                                           //Is the data in the tcp receive buffer to be analyzed bigger than 1 byte
                                           IF (#statReceive.trcvFct.dataLengthRest > 1) THEN
                                               //Yes --> get the telegram type in the 2nd byte
                                               #statReceive.tempTelegram.telegramType := #statReceive.trcvFct.data[#statReceive.trcvFct.dataOffset + 1];
                                           ELSE
                                               //No --> just one byte
                                               #statCopyNBytes := 1;
                                               #statReceive.tempTelegram.telegramType := 0;
                                           END_IF;

                                       ELSE
                                           //Already data in the temp. LCom header
                                           IF (#statReceive.tempTelegram.index = 1) THEN
                                               //Get the telegram type in the 1st byte
                                               #statReceive.tempTelegram.telegramType := #statReceive.trcvFct.data[#statReceive.trcvFct.dataOffset];
                                           ELSE
                                               //Get the telegram type in the 2nd byte
                                               #statReceive.tempTelegram.telegramType := #statReceive.trcvFct.data[#statReceive.trcvFct.dataOffset + 1];
                                           END_IF;
                                       END_IF;


                                       //---------------------------------------------------------------------
                                       //Build temp LCom header, if the telegram type is known
                                       //---------------------------------------------------------------------
                                       //Check if the telegram type is known
                                       IF (#statReceive.tempTelegram.telegramType > 0) THEN

                                           //Yes -->  telegram type is known
                                           CASE (#statReceive.tempTelegram.telegramType) OF
                                               1..3://Config telegram type 1,2,3
                                                   //LCom V2 (24 byte)
                                                   IF (#statReceive.tempTelegram.LComVersion = #HEADER_V2) THEN
                                                       IF ((24 - #statReceive.tempTelegram.index) < #statReceive.trcvFct.dataLengthRest) THEN
                                                           #statCopyNBytes := 24 - #statReceive.tempTelegram.index;
                                                       ELSE
                                                           #statCopyNBytes := #statReceive.trcvFct.dataLengthRest;
                                                       END_IF;
                                                   ELSE
                                                       //LCom V1 (16 byte)
                                                       IF ((16 - #statReceive.tempTelegram.index) < #statReceive.trcvFct.dataLengthRest) THEN
                                                           #statCopyNBytes := 16 - #statReceive.tempTelegram.index;
                                                       ELSE
                                                           #statCopyNBytes := #statReceive.trcvFct.dataLengthRest;
                                                       END_IF;
                                                   END_IF;
                                               5://Clock synchronization telegram type 5
                                                   //LCom V1 and V2 (10 byte)
                                                   IF ((10 - #statReceive.tempTelegram.index) < #statReceive.trcvFct.dataLengthRest) THEN
                                                       #statCopyNBytes := 10 - #statReceive.tempTelegram.index;
                                                   ELSE
                                                       #statCopyNBytes := #statReceive.trcvFct.dataLengthRest;
                                                   END_IF;
                                               10://Data telegram type 10
                                                   //LCom V2 (20 byte)
                                                   IF (#statReceive.tempTelegram.LComVersion = #HEADER_V2) THEN
                                                       IF ((20 - #statReceive.tempTelegram.index) < #statReceive.trcvFct.dataLengthRest) THEN
                                                           #statCopyNBytes := 20 - #statReceive.tempTelegram.index;
                                                       ELSE
                                                           #statCopyNBytes := #statReceive.trcvFct.dataLengthRest;
                                                       END_IF;
                                                   ELSE
                                                       //LCom V1 (12 byte)
                                                       IF ((12 - #statReceive.tempTelegram.index) < #statReceive.trcvFct.dataLengthRest) THEN
                                                           #statCopyNBytes := 12 - #statReceive.tempTelegram.index;
                                                       ELSE
                                                           #statCopyNBytes := #statReceive.trcvFct.dataLengthRest;
                                                       END_IF;
                                                   END_IF;
                                               20://Close connection telegram type 20
                                                   //LCom V1 (2 byte)
                                                   IF ((2 - #statReceive.tempTelegram.index) < #statReceive.trcvFct.dataLengthRest) THEN
                                                       #statCopyNBytes := 2 - #statReceive.tempTelegram.index;
                                                   ELSE
                                                       #statCopyNBytes := #statReceive.trcvFct.dataLengthRest;
                                                   END_IF;
                                               ELSE
                                                   //Write diagnostics
                                                   #statDiag.bufferIndex := #statDiag.bufferIndex + 1;
                                                   #statDiag.buffer[#statDiag.bufferIndex].status := #ERR_WRONG_TELEGRAM_ID;
                                                   #statDiag.buffer[#statDiag.bufferIndex].subFunctionErrorID := 16#0000;
                                                   #statDiag.buffer[#statDiag.bufferIndex].additionalValue1 := #statReceive.tempTelegram.telegramType;
                                                   #statDiag.buffer[#statDiag.bufferIndex].additionalValue2 := 0.0;
                                                   #statDiag.buffer[#statDiag.bufferIndex].additionalValue3 := 0.0;
                                                   #statDiag.buffer[#statDiag.bufferIndex].additionalValue4 := T#0ms;

                                                   #statState.connection := #CLOSE_CONNECTION;
                                                   GOTO diag;
                                           END_CASE;
                                       ELSE
                                           ;//No --> telegram type is zero
                                       END_IF;

                                       //Copy data into the temp. LCom header
                                       #statRet := MOVE_BLK_VARIANT(SRC := #statReceive.trcvFct.data, COUNT := #statCopyNBytes, SRC_INDEX := UDINT_TO_DINT(#statReceive.trcvFct.dataOffset), DEST_INDEX := #statReceive.tempTelegram.index, DEST => #statReceive.tempTelegram.data);
                                       //Calculate index in the temp. LCom header buffer
                                       #statReceive.tempTelegram.index := #statReceive.tempTelegram.index + UDINT_TO_USINT(#statCopyNBytes);
                                       //Calculate offset in the tcp receive buffer
                                       #statReceive.trcvFct.dataOffset := #statReceive.trcvFct.dataOffset + #statCopyNBytes;

                                       //Is local LCom version equal to partner LCom version ?
                                       IF (#statActualLocalLComVersion <> #statReceive.tempTelegram.LComVersion) THEN
                                           #statConnectAttempts := #statConnectAttempts + 1;
                                           //Write diagnostics
                                           #statDiag.bufferIndex := #statDiag.bufferIndex + 1;
                                           #statDiag.buffer[#statDiag.bufferIndex].status := #ERR_WRONG_HEADER;
                                           #statDiag.buffer[#statDiag.bufferIndex].subFunctionErrorID := 16#0000;
                                           #statDiag.buffer[#statDiag.bufferIndex].additionalValue1 := #statReceive.tempTelegram.LComVersion;
                                           #statDiag.buffer[#statDiag.bufferIndex].additionalValue2 := #statActualLocalLComVersion;
                                           #statDiag.buffer[#statDiag.bufferIndex].additionalValue3 := 0.0;
                                           #statDiag.buffer[#statDiag.bufferIndex].additionalValue4 := T#0ms;

                                           #statState.connection := #CLOSE_CONNECTION;
                                           GOTO diag;
                                       ELSE
                                           ;//local LCom version and partner LCom versions are equal
                                           #diagnostics.statistics.activeLComVersion := #statActualLocalLComVersion;
                                       END_IF;
                                   END_IF;//End: There is data expected without LCom header

                                   //---------------------------------------------------------------------
                                   //Interpret temp LCom header
                                   //---------------------------------------------------------------------
                                   IF (((#statReceive.tempTelegram.LComVersion = #HEADER_V1)//LCom V1
                                       AND//1,2,3 = 16 Byte
                                       ((#statReceive.tempTelegram.telegramType <= 3 AND #statReceive.tempTelegram.index = 16)
                                       OR//5 = 10 Byte
                                       (#statReceive.tempTelegram.telegramType = 5 AND #statReceive.tempTelegram.index = 10)
                                       OR//10 = 12 Byte
                                       (#statReceive.tempTelegram.telegramType = 10 AND #statReceive.tempTelegram.index = 12)
                                       OR//20 = 2 Byte
                                       (#statReceive.tempTelegram.telegramType = 20 AND #statReceive.tempTelegram.index = 2)))
                                       OR
                                       ((#statReceive.tempTelegram.LComVersion = #HEADER_V2)//LCom V2
                                       AND//1,2,3 = 24 Byte
                                       ((#statReceive.tempTelegram.telegramType <= 3 AND #statReceive.tempTelegram.index = 24)
                                       OR//5 = 10 Byte
                                       (#statReceive.tempTelegram.telegramType = 5 AND #statReceive.tempTelegram.index = 10)
                                       OR//10 = 20 Byte
                                       (#statReceive.tempTelegram.telegramType = 10 AND #statReceive.tempTelegram.index = 20)))
                                       OR
                                       (#statState.comReceiver = #DATA_EXPECTED))
                                   THEN

                                       CASE #statReceive.tempTelegram.telegramType OF

                                           10://Telegram type 10

                                               //Data expected without LCom header ?
                                               IF (#statState.comReceiver = #DATA_EXPECTED) THEN
                                                   //Yes --> LCom header from data telegram is already interpreted
                                                   //#receive.dataTelegram.messageOffset and #receive.dataTelegram.acPackageLength is known
                                                   //Calculate the bytes which have to be copied into FB.receiveData
                                                   IF (#statReceive.userData.offset + #statReceive.trcvFct.dataLengthRest) > (#statReceive.dataTelegram.messageOffset + #statReceive.dataTelegram.actPackageLength) THEN
                                                       //Copy just the missing bytes from the actual LCom package
                                                       #statCopyNBytes := ((#statReceive.dataTelegram.messageOffset + #statReceive.dataTelegram.actPackageLength) - #statReceive.userData.offset);
                                                   ELSE
                                                       //Copy all bytes which are still in the tcp receive buffer
                                                       #statCopyNBytes := #statReceive.trcvFct.dataLengthRest;
                                                   END_IF;
                                                   //Set SEND acknowledge message offset
                                                   #statSend.dataTelegram.ackMessageOffset := #statSend.dataTelegram.ackMessageOffset + #statCopyNBytes;
                                               ELSE
                                                   //Reset index, so a new temp. LCom header can be build
                                                   #statReceive.tempTelegram.index := 0;
                                                   #statReceive.numberOfLComHeader := #statReceive.numberOfLComHeader + 1;

                                                   //LComVersion
                                                   #statReceive.dataTelegram.LComVersion := #statReceive.tempTelegram.data[0];
                                                   //Telegram type
                                                   #statReceive.dataTelegram.telegramType := #statReceive.tempTelegram.data[1];
                                                   //Message counter
                                                   #statReceive.dataTelegram.messageCounter := #statReceive.tempTelegram.data[2];
                                                   //Acknowledge message counter
                                                   #statReceive.dataTelegram.ackMessageCounter := #statReceive.tempTelegram.data[3];

                                                   //LCom V2
                                                   IF (#statActualLocalLComVersion = #HEADER_V2) THEN
                                                       //Get tem. total message length
                                                       #tempDWord.%B3 := #statReceive.tempTelegram.data[16];
                                                       #tempDWord.%B2 := #statReceive.tempTelegram.data[17];
                                                       #tempDWord.%B1 := #statReceive.tempTelegram.data[18];
                                                       #tempDWord.%B0 := #statReceive.tempTelegram.data[19];

                                                       //Acknowledge message offset
                                                       #statReceive.dataTelegram.ackMessageOffset.%B3 := #statReceive.tempTelegram.data[8];
                                                       #statReceive.dataTelegram.ackMessageOffset.%B2 := #statReceive.tempTelegram.data[9];
                                                       #statReceive.dataTelegram.ackMessageOffset.%B1 := #statReceive.tempTelegram.data[10];
                                                       #statReceive.dataTelegram.ackMessageOffset.%B0 := #statReceive.tempTelegram.data[11];

                                                       //Is it an acknowledge telegram ?
                                                       IF (#tempDWord = 16#0000) THEN
                                                           //Acknowledge telegram
                                                           #statState.comReceiver := #ACK_TELEGRAM;
                                                       ELSE
                                                           //Is no acknowledge telegram
                                                           //Message offset
                                                           #statReceive.dataTelegram.messageOffset.%B3 := #statReceive.tempTelegram.data[4];
                                                           #statReceive.dataTelegram.messageOffset.%B2 := #statReceive.tempTelegram.data[5];
                                                           #statReceive.dataTelegram.messageOffset.%B1 := #statReceive.tempTelegram.data[6];
                                                           #statReceive.dataTelegram.messageOffset.%B0 := #statReceive.tempTelegram.data[7];
                                                           //Actual package length
                                                           #statReceive.dataTelegram.actPackageLength.%B3 := #statReceive.tempTelegram.data[12];
                                                           #statReceive.dataTelegram.actPackageLength.%B2 := #statReceive.tempTelegram.data[13];
                                                           #statReceive.dataTelegram.actPackageLength.%B1 := #statReceive.tempTelegram.data[14];
                                                           #statReceive.dataTelegram.actPackageLength.%B0 := #statReceive.tempTelegram.data[15];
                                                           //Total message length
                                                           #statReceive.dataTelegram.totalMessageLength := #tempDWord;
                                                       END_IF;
                                                   ELSE
                                                       //LCom V1
                                                       //Get temp. total message length
                                                       #tempDWord.%B1 := #statReceive.tempTelegram.data[10];
                                                       #tempDWord.%B0 := #statReceive.tempTelegram.data[11];

                                                       //Acknowledge message offset
                                                       #statReceive.dataTelegram.ackMessageOffset.%B1 := #statReceive.tempTelegram.data[6];
                                                       #statReceive.dataTelegram.ackMessageOffset.%B0 := #statReceive.tempTelegram.data[7];

                                                       //Is it an acknowledge telegram ?
                                                       IF (#tempDWord = 16#0000) THEN
                                                           //Acknowledge telegram
                                                           #statState.comReceiver := #ACK_TELEGRAM;
                                                       ELSE
                                                           //Is no acknowledge telegram
                                                           //Message offset
                                                           #statReceive.dataTelegram.messageOffset.%B1 := #statReceive.tempTelegram.data[4];
                                                           #statReceive.dataTelegram.messageOffset.%B0 := #statReceive.tempTelegram.data[5];
                                                           //Actual package length
                                                           #statReceive.dataTelegram.actPackageLength.%B1 := #statReceive.tempTelegram.data[8];
                                                           #statReceive.dataTelegram.actPackageLength.%B0 := #statReceive.tempTelegram.data[9];
                                                           //Total message length
                                                           #statReceive.dataTelegram.totalMessageLength := #tempDWord;
                                                       END_IF;
                                                   END_IF;

                                                   //Set SEND acknowledge message offset
                                                   #statSend.dataTelegram.ackMessageCounter := #statReceive.dataTelegram.messageCounter;

                                                   //Check if the LCom package, which was sent before is acknowledged ?
                                                   IF ((#statSend.numberOfLComPackage = 1)//One package was sent
                                                       AND
                                                       ((#statSend.expectedAck.package1.offset = #statReceive.dataTelegram.ackMessageOffset)
                                                       AND
                                                       (#statSend.dataTelegram.messageCounter = #statReceive.dataTelegram.ackMessageCounter)))
                                                   THEN
                                                       //Acknowledgement for the package x.1
                                                       #statSend.numberOfLComPackage := 0;
                                                       //Stop acknowledge timer for the 1st package
                                                       #instExpectedAckPackage1(IN := FALSE,
                                                                                PT := #diagnostics.localConfig.sender.ackTimeout);
                                                   ELSIF ((#statSend.dataTelegram.messageCounter = #statReceive.dataTelegram.ackMessageCounter)
                                                       OR
                                                       (#statSend.dataTelegram.messageCounter - 1 = #statReceive.dataTelegram.ackMessageCounter)
                                                       OR
                                                       (#diagnostics.statistics.maxMsgSendingTime = T#0ms))//Workaround: S7 Controller does not start with correct ack. message counter
                                                   THEN
                                                       ;
                                                   ELSE
                                                       //Write diagnostics
                                                       #statDiag.bufferIndex := #statDiag.bufferIndex + 1;
                                                       #statDiag.buffer[#statDiag.bufferIndex].status := #ERR_ACK_MESSAGE_NUMBER;
                                                       #statDiag.buffer[#statDiag.bufferIndex].subFunctionErrorID := 16#0000;
                                                       #statDiag.buffer[#statDiag.bufferIndex].additionalValue1 := #statReceive.dataTelegram.messageCounter;
                                                       #statDiag.buffer[#statDiag.bufferIndex].additionalValue2 := #statSend.dataTelegram.messageCounter;
                                                       #statDiag.buffer[#statDiag.bufferIndex].additionalValue3 := 0.0;
                                                       #statDiag.buffer[#statDiag.bufferIndex].additionalValue4 := T#0ms;

                                                       #statState.connection := #CLOSE_CONNECTION;
                                                       GOTO diag;
                                                   END_IF;


                                                   //Is the 1st LCom package received and nothing is copied into FB.receiveData so far ?
                                                   IF ((#statReceive.userData.totalLength = 0)
                                                       AND
                                                       (#statReceive.dataTelegram.messageOffset = 0)
                                                       AND
                                                       (#statState.comReceiver <> #ACK_TELEGRAM))
                                                   THEN
                                                       //Store the 1st received telegram with the total receive length
                                                       #statReceive.userData.totalLength := #statReceive.dataTelegram.totalMessageLength;
                                                       //Reset the acknowledged message offset
                                                       #statSend.dataTelegram.ackMessageOffset := 0;

                                                       //Start message receiving timer
                                                       #instMsgReceivingTimer(IN := TRUE,
                                                                              PT := T#+24d20h31m23s647ms);
                                                   ELSE
                                                       ;//In receiving process or acknowledge telegram
                                                   END_IF;

                                                   //Is the data telegram a acknowledge telegram ?
                                                   IF (#statState.comReceiver = #ACK_TELEGRAM)
                                                   THEN
                                                       //Yes --> Acknowledge telegram, no bytes have to be copied
                                                       #statCopyNBytes := 0;
                                                   ELSIF ((#diagnostics.statistics.activeLComVersion = #HEADER_V1)
                                                       AND
                                                       ((#statReceive.userData.offset + (#statReceive.trcvFct.dataLengthRest - 12)) > (#statReceive.dataTelegram.messageOffset + #statReceive.dataTelegram.actPackageLength)))
                                                   THEN//No --> The data to be analyzed in the tcp receive buffer is bigger than the complete message

                                                       //Do not copy all data from the tcp receive buffer, only the rest data from the LCom package
                                                       #statCopyNBytes := ((#statReceive.dataTelegram.messageOffset + #statReceive.dataTelegram.actPackageLength) - #statReceive.userData.offset);
                                                       //Calculate acknowledge message offset which has to be sent to the partner
                                                       #statSend.dataTelegram.ackMessageOffset := #statSend.dataTelegram.ackMessageOffset + #statCopyNBytes;
                                                   ELSIF ((#diagnostics.statistics.activeLComVersion = #HEADER_V2)
                                                       AND
                                                       ((#statReceive.userData.offset + (#statReceive.trcvFct.dataLengthRest - 24)) > (#statReceive.dataTelegram.messageOffset + #statReceive.dataTelegram.actPackageLength)))
                                                   THEN//No --> The data to be analyzed in the tcp receive buffer is bigger than the complete message

                                                       //Copy not all data from the tcp receive buffer, only the rest data from the LCom package
                                                       #statCopyNBytes := ((#statReceive.dataTelegram.messageOffset + #statReceive.dataTelegram.actPackageLength) - #statReceive.userData.offset);
                                                       //Calculate acknowledge message offset which have to be sent to the partner
                                                       #statSend.dataTelegram.ackMessageOffset := #statSend.dataTelegram.ackMessageOffset + #statCopyNBytes;
                                                   ELSE
                                                       //Copy just the rest of data from the tcp receive buffer
                                                       IF #diagnostics.statistics.activeLComVersion = #HEADER_V1 THEN
                                                           #statCopyNBytes := #statReceive.trcvFct.dataLengthRest - 12;
                                                       ELSE
                                                           #statCopyNBytes := #statReceive.trcvFct.dataLengthRest - 20;
                                                       END_IF;
                                                       //Calculate acknowledge message offset which have to be sent to the partner
                                                       #statSend.dataTelegram.ackMessageOffset := #statSend.dataTelegram.ackMessageOffset + #statCopyNBytes;
                                                   END_IF;

                                               END_IF;

                                               //Copy data to FB.receiveBuffer
                                               #statRet := MOVE_BLK_VARIANT(SRC := #statReceive.trcvFct.data, COUNT := #statCopyNBytes, SRC_INDEX := UDINT_TO_DINT(#statReceive.trcvFct.dataOffset), DEST_INDEX := UDINT_TO_DINT(#statReceive.userData.offset), DEST => #receiveBuffer);
                                               //Calculate offset in the FB.#receiveBuffer
                                               #statReceive.userData.offset := #statReceive.userData.offset + #statCopyNBytes;
                                               //Calculate offset in the tcp receive buffer
                                               #statReceive.trcvFct.dataOffset := #statReceive.trcvFct.dataOffset + #statCopyNBytes;

                                               //---------------------------------------------------------------------
                                               //Is complete LCom message acknowledged which was sent ?
                                               //---------------------------------------------------------------------
                                               IF ((#statSend.userData.offset = #statReceive.dataTelegram.ackMessageOffset)
                                                   AND
                                                   (#statReceive.dataTelegram.ackMessageCounter = #statSend.dataTelegram.messageCounter)
                                                   AND
                                                   #statState.comSender = #SEND_NO_DATA)
                                               THEN
                                                   //Yes --> Complete LCom message is acknowledged
                                                   #sending := #statSending := FALSE;

                                                   //Statistic --> Increase number of sent user messages
                                                   #diagnostics.statistics.numberOfSentMessages := #diagnostics.statistics.numberOfSentMessages + 1;

                                                   //Get message sending time [ms]
                                                   #instMsgSendingTimer(IN := TRUE,
                                                                        PT := T#+24d20h31m23s647ms);

                                                   //Statistic --> Compare max. message sending time
                                                   IF (#instMsgSendingTimer.ET > #diagnostics.statistics.maxMsgSendingTime) THEN
                                                       #diagnostics.statistics.maxMsgSendingTime := #instMsgSendingTimer.ET;
                                                   ELSE
                                                       ;//Actual sending time is smaller
                                                   END_IF;

                                                   //Statistic --> Calculate average of message sending time [ms)]
                                                   #diagnostics.statistics.avgMsgSendingTime := (((#diagnostics.statistics.avgMsgSendingTime * 19) + UDINT_TO_REAL((TIME_TO_UDINT(#instMsgSendingTimer.ET)))) / 20);

                                                   //Stop message sending timer
                                                   #instMsgSendingTimer(IN := FALSE,
                                                                        PT := T#+24d20h31m23s647ms);

                                                   //Initialize values, for next send request
                                                   #statSend.userData.offset := 0;
                                                   #statSend.dataTelegram.messageOffset := 0;
                                                   #statSend.dataTelegram.totalMessageLength := 0;
                                               ELSE
                                                   ;//Complete LCom message is not acknowledged yet
                                               END_IF;//End: Is complete Lcom message acknowledged, which was sent ?


                                               //---------------------------------------------------------------------
                                               //Build acknowledge telegram
                                               //---------------------------------------------------------------------

                                               //Assume always that an LCom package is expected
                                               #statState.comReceiver := #EXPECTED;

                                               //---------------------------------------------------------------------
                                               //Has the complete LCom package been received (1 Byte ... 4 Kilobyte) ?
                                               //---------------------------------------------------------------------
                                               IF (#statReceive.userData.offset = 0) THEN
                                                   ;//Do nothing
                                               ELSIF (#statReceive.userData.offset = (#statReceive.dataTelegram.messageOffset + #statReceive.dataTelegram.actPackageLength))
                                               THEN//Yes --> Complete LCom package has been received (1 Byte ... 4k Byte)

                                                   //Still in sending process and LCom package sent is not acknowledged yet ?
                                                   //Select LCom V1 or V2; now one LCom package is sent and must be acknowledged
                                                   IF ((#statSending = TRUE)
                                                       AND
                                                       (#statSend.numberOfLComPackage = 0)
                                                       AND
                                                       ((#statActualLocalLComVersion = #HEADER_V1)
                                                       OR
                                                       (#statActualLocalLComVersion = #HEADER_V2)))
                                                   THEN
                                                       ;//Build no acknowledge telegram 10
                                                   ELSE
                                                       //Build acknowledge telegram 10
                                                       #statSend.tsendFct.data[#statSend.tsendFct.dataOffset] := #statSend.dataTelegram.LComVersion;
                                                       #statSend.tsendFct.data[#statSend.tsendFct.dataOffset + 1] := #statSend.dataTelegram.telegramType;
                                                       #statSend.tsendFct.data[#statSend.tsendFct.dataOffset + 2] := #statSend.dataTelegram.messageCounter;
                                                       #statSend.tsendFct.data[#statSend.tsendFct.dataOffset + 3] := #statSend.dataTelegram.ackMessageCounter;
                                                       //Message offset
                                                       #statSend.tsendFct.data[#statSend.tsendFct.dataOffset + 4] := 16#00;
                                                       #statSend.tsendFct.data[#statSend.tsendFct.dataOffset + 5] := 16#00;
                                                       #statSend.tsendFct.data[#statSend.tsendFct.dataOffset + 6] := 16#00;
                                                       #statSend.tsendFct.data[#statSend.tsendFct.dataOffset + 7] := 16#00;
                                                       //Acknowledge message offset
                                                       #statSend.tsendFct.data[#statSend.tsendFct.dataOffset + 8] := #statSend.dataTelegram.ackMessageOffset.%B3;
                                                       #statSend.tsendFct.data[#statSend.tsendFct.dataOffset + 9] := #statSend.dataTelegram.ackMessageOffset.%B2;
                                                       #statSend.tsendFct.data[#statSend.tsendFct.dataOffset + 10] := #statSend.dataTelegram.ackMessageOffset.%B1;
                                                       #statSend.tsendFct.data[#statSend.tsendFct.dataOffset + 11] := #statSend.dataTelegram.ackMessageOffset.%B0;
                                                       //Actual package length
                                                       #statSend.tsendFct.data[#statSend.tsendFct.dataOffset + 12] := 16#00;
                                                       #statSend.tsendFct.data[#statSend.tsendFct.dataOffset + 13] := 16#00;
                                                       #statSend.tsendFct.data[#statSend.tsendFct.dataOffset + 14] := 16#00;
                                                       #statSend.tsendFct.data[#statSend.tsendFct.dataOffset + 15] := 16#00;
                                                       //Total message length
                                                       #statSend.tsendFct.data[#statSend.tsendFct.dataOffset + 16] := 16#00;
                                                       #statSend.tsendFct.data[#statSend.tsendFct.dataOffset + 17] := 16#00;
                                                       #statSend.tsendFct.data[#statSend.tsendFct.dataOffset + 18] := 16#00;
                                                       #statSend.tsendFct.data[#statSend.tsendFct.dataOffset + 19] := 16#00;

                                                       //LCom V2
                                                       IF (#statActualLocalLComVersion = #HEADER_V2) THEN
                                                           //Calculate offset in the tcp send buffer
                                                           #statSend.tsendFct.dataOffset := #statSend.tsendFct.dataOffset + 20;
                                                       ELSE
                                                           //LCom V1
                                                           //Acknowledge message offset
                                                           #statSend.tsendFct.data[#statSend.tsendFct.dataOffset + 6] := #statSend.dataTelegram.ackMessageOffset.%B1;
                                                           #statSend.tsendFct.data[#statSend.tsendFct.dataOffset + 7] := #statSend.dataTelegram.ackMessageOffset.%B0;
                                                           //Actual package length
                                                           #statSend.tsendFct.data[#statSend.tsendFct.dataOffset + 8] := 16#00;
                                                           #statSend.tsendFct.data[#statSend.tsendFct.dataOffset + 9] := 16#00;
                                                           //Total message length
                                                           #statSend.tsendFct.data[#statSend.tsendFct.dataOffset + 10] := 16#00;
                                                           #statSend.tsendFct.data[#statSend.tsendFct.dataOffset + 11] := 16#00;
                                                           //Calculate offset in the tcp send buffer
                                                           #statSend.tsendFct.dataOffset := #statSend.tsendFct.dataOffset + 12;
                                                       END_IF;
                                                       //Set sender state
                                                       #statState.sender := #SEND_CONFIG;
                                                   END_IF;


                                                   //---------------------------------------------------------------------
                                                   //Is the complete LCom message received (1 Byte ... 4 Gigabyte) ?
                                                   //---------------------------------------------------------------------
                                                   IF (#statReceive.userData.offset = #statReceive.dataTelegram.totalMessageLength) THEN
                                                       //Yes --> Set FB outputs
                                                       #dataReceived := #statDataReceived := TRUE;
                                                       #receivedDataLength := #statReceive.dataTelegram.totalMessageLength;
                                                       //Initialize values, for next receive request
                                                       #statReceive.userData.totalLength := 0;
                                                       #statReceive.userData.offset := 0;

                                                       //Statistic --> Increase number of received user messages
                                                       #diagnostics.statistics.numberOfReceivedMessages := #diagnostics.statistics.numberOfReceivedMessages + 1;

                                                       //Get message receiving time [ms]
                                                       #instMsgReceivingTimer(IN := TRUE,
                                                                              PT := T#+24d20h31m23s647ms);

                                                       //Statistic --> Compare max. message receiving time
                                                       IF (#instMsgReceivingTimer.ET > #diagnostics.statistics.maxMsgReceivingTime) THEN
                                                           #diagnostics.statistics.maxMsgReceivingTime := #instMsgReceivingTimer.ET;
                                                       ELSE
                                                           ;//Actual receiving time is smaller
                                                       END_IF;

                                                       //Statistic --> Calculate average of message receiving time [ms]
                                                       #diagnostics.statistics.avgMsgReceivingTime := (((#diagnostics.statistics.avgMsgReceivingTime * 19) + UDINT_TO_REAL((TIME_TO_UDINT(#instMsgReceivingTimer.ET)))) / 20);

                                                       //Stop message receiving timer
                                                       #instMsgReceivingTimer(IN := FALSE,
                                                                              PT := T#+24d20h31m23s647ms);


                                                       //Get received messages cycle time [ms]
                                                       #instReceiveMsgCycle(IN := TRUE,
                                                                            PT := T#+24d20h31m23s647ms);

                                                       //Statistic --> Compare max. received messages cycle time
                                                       IF (#instReceiveMsgCycle.ET > #diagnostics.statistics.maxReceiveMsgCycle) THEN
                                                           #diagnostics.statistics.maxReceiveMsgCycle := #instReceiveMsgCycle.ET;
                                                       ELSE
                                                           ;//Actual receiving time is smaller
                                                       END_IF;

                                                       //Statistic --> Check receive messages cycle time violations (receive cycle time >= 110%)
                                                       IF (#instReceiveMsgCycle.ET > (#diagnostics.partnerConfig.sender.cycleTime + (#diagnostics.partnerConfig.sender.cycleTime / 10))) THEN
                                                           #diagnostics.statistics.totalReceiveCycleViolations := #diagnostics.statistics.totalReceiveCycleViolations + 1;
                                                       ELSE
                                                           ;//Receive messages cycle time is smaller
                                                       END_IF;

                                                       //Statistic --> calculate average of receive messages cycle time [ms]
                                                       #diagnostics.statistics.avgReceiveMsgCycle := (((#diagnostics.statistics.avgReceiveMsgCycle * 19) + UDINT_TO_REAL((TIME_TO_UDINT(#instReceiveMsgCycle.ET)))) / 20);

                                                       //Stop received message timer
                                                       #instReceiveMsgCycle(IN := false,
                                                                            PT := T#+24d20h31m23s647ms);

                                                       //Start received message timer
                                                       #instReceiveMsgCycle(IN := TRUE,
                                                                            PT := T#+24d20h31m23s647ms);

                                                   ELSE
                                                       //No --> Still more LCom package expected
                                                       #statState.comReceiver := #EXPECTED;
                                                   END_IF;//End: Is the complete LCom message received (1 Byte ... 4 Gigabyte)
                                               ELSE
                                                   //Data without LCom Header expected
                                                   #statState.comReceiver := #DATA_EXPECTED;
                                               END_IF;//Is the complete LCom package received (1 Byte ... 4 Kilobyte)

                                           3://Telegram type 3

                                               //Reset index, so a new temp. LCom header can be built
                                               #statReceive.tempTelegram.index := 0;
                                               #statReceive.numberOfLComHeader := #statReceive.numberOfLComHeader + 1;

                                               //Partner information is already known in the diagnostic structure
                                               IF (#diagnostics.partnerConfig.connnection.lifeSignCycleTime = T#0ms) THEN
                                                   //No --> Get diagnostics information
                                                   //LCom V2
                                                   IF (#statActualLocalLComVersion = #HEADER_V2) THEN
                                                       //UsesTimeStamp
                                                       #diagnostics.partnerConfig.timeSync.usePartnerTimestamps := BYTE_TO_BOOL(#statReceive.tempTelegram.data[2]);
                                                       //SendModeSyncTime
                                                       #diagnostics.partnerConfig.timeSync.sendMode := #statReceive.tempTelegram.data[3];
                                                       //LifeSignCycle
                                                       #tempDWord.%B3 := #statReceive.tempTelegram.data[4];
                                                       #tempDWord.%B2 := #statReceive.tempTelegram.data[5];
                                                       #tempDWord.%B1 := #statReceive.tempTelegram.data[6];
                                                       #tempDWord.%B0 := #statReceive.tempTelegram.data[7];
                                                       #statReceive.configTelegramV2.lifeSignCycle := DWORD_TO_TIME(#tempDWord);
                                                       #diagnostics.partnerConfig.connnection.lifeSignCycleTime := #statReceive.configTelegramV2.lifeSignCycle;
                                                       //Sender cycleTime
                                                       #tempDWord.%B3 := #statReceive.tempTelegram.data[8];
                                                       #tempDWord.%B2 := #statReceive.tempTelegram.data[9];
                                                       #tempDWord.%B1 := #statReceive.tempTelegram.data[10];
                                                       #tempDWord.%B0 := #statReceive.tempTelegram.data[11];
                                                       #statReceive.configTelegramV2.cycleTime := DWORD_TO_TIME(#tempDWord);
                                                       #diagnostics.partnerConfig.sender.cycleTime := #statReceive.configTelegramV2.cycleTime;
                                                       //Sender ackTimeOut
                                                       #tempDWord.%B3 := #statReceive.tempTelegram.data[12];
                                                       #tempDWord.%B2 := #statReceive.tempTelegram.data[13];
                                                       #tempDWord.%B1 := #statReceive.tempTelegram.data[14];
                                                       #tempDWord.%B0 := #statReceive.tempTelegram.data[15];
                                                       #statReceive.configTelegramV2.ackTimeOut := DWORD_TO_TIME(#tempDWord);
                                                       #diagnostics.partnerConfig.sender.ackTimeout := #statReceive.configTelegramV2.ackTimeOut;
                                                       //MaxSendDataLength
                                                       #tempDWord.%B3 := #statReceive.tempTelegram.data[16];
                                                       #tempDWord.%B2 := #statReceive.tempTelegram.data[17];
                                                       #tempDWord.%B1 := #statReceive.tempTelegram.data[18];
                                                       #tempDWord.%B0 := #statReceive.tempTelegram.data[19];
                                                       #statReceive.configTelegramV2.maxSendDataLength := #tempDWord;
                                                       #diagnostics.partnerConfig.sizeOfSendBuffer := #statReceive.configTelegramV2.maxSendDataLength;
                                                       //MaxReceiveDataLength
                                                       #tempDWord.%B3 := #statReceive.tempTelegram.data[20];
                                                       #tempDWord.%B2 := #statReceive.tempTelegram.data[21];
                                                       #tempDWord.%B1 := #statReceive.tempTelegram.data[22];
                                                       #tempDWord.%B0 := #statReceive.tempTelegram.data[23];
                                                       #statReceive.configTelegramV2.maxReceiveDataLength := #tempDWord;
                                                       #diagnostics.partnerConfig.sizeOfReceiveBuffer := #statReceive.configTelegramV2.maxReceiveDataLength;
                                                   ELSE
                                                       //LCom V1
                                                       //LifeSignCycle
                                                       #statReceive.configTelegramV1.lifeSignCycle.%B1 := #statReceive.tempTelegram.data[8];
                                                       #statReceive.configTelegramV1.lifeSignCycle.%B0 := #statReceive.tempTelegram.data[9];
                                                       #diagnostics.partnerConfig.connnection.lifeSignCycleTime := UINT_TO_TIME(#statReceive.configTelegramV1.lifeSignCycle);
                                                       //MaxSendDataLength
                                                       #statReceive.configTelegramV1.maxSendDataLength.%B1 := #statReceive.tempTelegram.data[12];
                                                       #statReceive.configTelegramV1.maxSendDataLength.%B0 := #statReceive.tempTelegram.data[13];
                                                       #diagnostics.partnerConfig.sizeOfSendBuffer := #statReceive.configTelegramV1.maxSendDataLength;
                                                       //MaxReceiveDataLength
                                                       #statReceive.configTelegramV1.maxReceiveDataLength.%B1 := #statReceive.tempTelegram.data[14];
                                                       #statReceive.configTelegramV1.maxReceiveDataLength.%B0 := #statReceive.tempTelegram.data[15];
                                                       #diagnostics.partnerConfig.sizeOfReceiveBuffer := #statReceive.configTelegramV1.maxReceiveDataLength;
                                                       //UsesTimeStamp
                                                       #diagnostics.partnerConfig.timeSync.usePartnerTimestamps := BYTE_TO_BOOL(#statReceive.tempTelegram.data[10]);
                                                       //SendModeSyncTime
                                                       #diagnostics.partnerConfig.timeSync.sendMode := #statReceive.tempTelegram.data[11];
                                                   END_IF;
                                               END_IF;

                                           1://Telegram type 1

                                               //Reset index, so a new temp. LCom header can be built
                                               #statReceive.tempTelegram.index := 0;
                                               #statReceive.numberOfLComHeader := #statReceive.numberOfLComHeader + 1;

                                               //LCom V1
                                               //LifeSignCycle
                                               #statReceive.configTelegramV1.lifeSignCycle.%B1 := #statReceive.tempTelegram.data[8];
                                               #statReceive.configTelegramV1.lifeSignCycle.%B0 := #statReceive.tempTelegram.data[9];
                                               #diagnostics.partnerConfig.connnection.lifeSignCycleTime := UINT_TO_TIME(#statReceive.configTelegramV1.lifeSignCycle);
                                               //Receiver cycleTime from receiver
                                               #statReceive.configTelegramV1.cycleTime.%B1 := #statReceive.tempTelegram.data[4];
                                               #statReceive.configTelegramV1.cycleTime.%B0 := #statReceive.tempTelegram.data[5];
                                               //Receiver ackTimeOut from receiver
                                               #statReceive.configTelegramV1.ackTimeOut.%B1 := #statReceive.tempTelegram.data[6];
                                               #statReceive.configTelegramV1.ackTimeOut.%B0 := #statReceive.tempTelegram.data[7];

                                               //Are receive cycle time and current sender cycle time and receive ackTimeOut and current sender ackTimeOut equal ?
                                               IF ((#statReceive.configTelegramV1.cycleTime = (TIME_TO_UINT(#diagnostics.localConfig.sender.cycleTime)))
                                                   AND
                                                   (#statReceive.configTelegramV1.ackTimeOut = (TIME_TO_UINT(#diagnostics.localConfig.sender.ackTimeout))))
                                               THEN
                                                   ;//Yes equal --> Set FB.#connected and diagnostics information
                                               ELSE
                                                   //Not equal --> Compare values and prioritize
                                                   //Compare cycle time
                                                   IF (#statReceive.configTelegramV1.cycleTime > (TIME_TO_UINT(#diagnostics.localConfig.sender.cycleTime))) THEN
                                                       #statSend.configTelegramV1.cycleTime := #statReceive.configTelegramV1.cycleTime;
                                                   ELSE
                                                       ;//Actual sender cycleTime is bigger than the received sender cycleTime
                                                   END_IF;

                                                   //Compare acknowledge timeout
                                                   IF (#statReceive.configTelegramV1.ackTimeOut > (TIME_TO_UINT(#diagnostics.localConfig.sender.ackTimeout))) THEN
                                                       #statSend.configTelegramV1.ackTimeOut := #statReceive.configTelegramV1.ackTimeOut;
                                                   ELSE
                                                       ;//Actual acknowledge timeout is bigger than the received sender acknowledge timeout
                                                   END_IF;

                                                   //Update diagnostics information
                                                   #diagnostics.localConfig.sender.cycleTime := UINT_TO_TIME(#statReceive.configTelegramV1.cycleTime);
                                                   #diagnostics.localConfig.sender.ackTimeout := UINT_TO_TIME(#statReceive.configTelegramV1.ackTimeOut);

                                                   //Send telegram 2
                                                   #statSend.tsendFct.data[#statSend.tsendFct.dataOffset] := #statSend.configTelegramV1.LComVersion;
                                                   #statSend.tsendFct.data[#statSend.tsendFct.dataOffset + 1] := 16#02;
                                                   #statSend.tsendFct.data[#statSend.tsendFct.dataOffset + 2] := #statSend.configTelegramV1.comMode;
                                                   #statSend.tsendFct.data[#statSend.tsendFct.dataOffset + 3] := #statSend.configTelegramV1.slidingWindow;
                                                   //Cycle time
                                                   #statSend.tsendFct.data[#statSend.tsendFct.dataOffset + 4] := #statSend.configTelegramV1.cycleTime.%B1;
                                                   #statSend.tsendFct.data[#statSend.tsendFct.dataOffset + 5] := #statSend.configTelegramV1.cycleTime.%B0;
                                                   //Acknowledge timeout
                                                   #statSend.tsendFct.data[#statSend.tsendFct.dataOffset + 6] := #statSend.configTelegramV1.ackTimeOut.%B1;
                                                   #statSend.tsendFct.data[#statSend.tsendFct.dataOffset + 7] := #statSend.configTelegramV1.ackTimeOut.%B0;
                                                   //LifeSignCycle
                                                   #statSend.tsendFct.data[#statSend.tsendFct.dataOffset + 8] := #statSend.configTelegramV1.lifeSignCycle.%B1;
                                                   #statSend.tsendFct.data[#statSend.tsendFct.dataOffset + 9] := #statSend.configTelegramV1.lifeSignCycle.%B0;
                                                   //Status
                                                   #statSend.tsendFct.data[#statSend.tsendFct.dataOffset + 10] := #statSend.configTelegramV1.status;
                                                   //SendModeSyncTime
                                                   #statSend.tsendFct.data[#statSend.tsendFct.dataOffset + 11] := #statSend.configTelegramV1.sendModeSyncTime;
                                                   //MaxSendDataLength
                                                   #statSend.tsendFct.data[#statSend.tsendFct.dataOffset + 12] := #statSend.configTelegramV1.maxSendDataLength.%B1;
                                                   #statSend.tsendFct.data[#statSend.tsendFct.dataOffset + 13] := #statSend.configTelegramV1.maxSendDataLength.%B0;
                                                   //MaxReceiveDataLength
                                                   #statSend.tsendFct.data[#statSend.tsendFct.dataOffset + 14] := #statSend.configTelegramV1.maxReceiveDataLength.%B1;
                                                   #statSend.tsendFct.data[#statSend.tsendFct.dataOffset + 15] := #statSend.configTelegramV1.maxReceiveDataLength.%B0;
                                                   //Calculate offset in the tcp send buffer
                                                   #statSend.tsendFct.dataOffset := #statSend.tsendFct.dataOffset + 16;
                                                   #statState.sender := #SEND_CONFIG;
                                               END_IF;

                                               //Set FB.#connected and #diagnostics information
                                               #connected := #statConnected := TRUE;
                                               #diagnostics.statistics.LComProtocolUsed := TRUE;
                                               #diagnostics.statistics.activeLComVersion := #HEADER_V1;
                                               //Write diagnostics
                                               #statDiag.bufferIndex := #statDiag.bufferIndex + 1;
                                               #statDiag.buffer[#statDiag.bufferIndex].status := #STATUS_CONNECTED_V1;
                                               #statDiag.buffer[#statDiag.bufferIndex].subFunctionErrorID := 16#0000;
                                               #statDiag.buffer[#statDiag.bufferIndex].additionalValue1 := 0.0;
                                               #statDiag.buffer[#statDiag.bufferIndex].additionalValue2 := 0.0;
                                               #statDiag.buffer[#statDiag.bufferIndex].additionalValue3 := 0.0;
                                               #statDiag.buffer[#statDiag.bufferIndex].additionalValue4 := T#0ms;

                                               #statState.cfgSender := #OPERATION;

                                               //MaxSendDataLength
                                               #statReceive.configTelegramV1.maxSendDataLength.%B1 := #statReceive.tempTelegram.data[12];
                                               #statReceive.configTelegramV1.maxSendDataLength.%B0 := #statReceive.tempTelegram.data[13];
                                               #diagnostics.partnerConfig.sizeOfSendBuffer := #statReceive.configTelegramV1.maxSendDataLength;
                                               //MaxReceiveDataLength
                                               #statReceive.configTelegramV1.maxReceiveDataLength.%B1 := #statReceive.tempTelegram.data[14];
                                               #statReceive.configTelegramV1.maxReceiveDataLength.%B0 := #statReceive.tempTelegram.data[15];
                                               #diagnostics.partnerConfig.sizeOfReceiveBuffer := #statReceive.configTelegramV1.maxReceiveDataLength;
                                               //UsesTimeStamp
                                               #diagnostics.partnerConfig.timeSync.usePartnerTimestamps := BYTE_TO_BOOL(#statReceive.tempTelegram.data[10]);
                                               //SendModeSyncTime
                                               #diagnostics.partnerConfig.timeSync.sendMode := #statReceive.tempTelegram.data[11];

                                               IF ((#diagnostics.localConfig.timeSync.usePartnerTimestamps
                                                   XOR
                                                   #diagnostics.partnerConfig.timeSync.usePartnerTimestamps)
                                                   AND
                                                   (#diagnostics.localConfig.timeSync.sendMode > 0
                                                   OR
                                                   #diagnostics.partnerConfig.timeSync.sendMode > 0))
                                               THEN
                                                   ;//One cpu does send timeSync information
                                               ELSE
                                                   //Write diagnostics
                                                   #statDiag.bufferIndex := #statDiag.bufferIndex + 1;
                                                   #statDiag.buffer[#statDiag.bufferIndex].status := #WARN_NO_TIME_SYNC;
                                                   #statDiag.buffer[#statDiag.bufferIndex].subFunctionErrorID := 16#0000;
                                                   #statDiag.buffer[#statDiag.bufferIndex].additionalValue1 := 0.0;
                                                   #statDiag.buffer[#statDiag.bufferIndex].additionalValue2 := 0.0;
                                                   #statDiag.buffer[#statDiag.bufferIndex].additionalValue3 := 0.0;
                                                   #statDiag.buffer[#statDiag.bufferIndex].additionalValue4 := T#0ms;
                                               END_IF;

                                           2://telegram type 2

                                               //Reset index, so a new temp. LCom header can be built
                                               #statReceive.tempTelegram.index := 0;
                                               #statReceive.numberOfLComHeader := #statReceive.numberOfLComHeader + 1;

                                               //LCom V2
                                               IF (#statActualLocalLComVersion = #HEADER_V2) THEN
                                                   //UsesTimeStamp
                                                   #diagnostics.partnerConfig.timeSync.usePartnerTimestamps := BYTE_TO_BOOL(#statReceive.tempTelegram.data[2]);
                                                   //SendModeSyncTime
                                                   #diagnostics.partnerConfig.timeSync.sendMode := #statReceive.tempTelegram.data[3];
                                                   //LifeSignCycle
                                                   #tempDWord.%B3 := #statReceive.tempTelegram.data[4];
                                                   #tempDWord.%B2 := #statReceive.tempTelegram.data[5];
                                                   #tempDWord.%B1 := #statReceive.tempTelegram.data[6];
                                                   #tempDWord.%B0 := #statReceive.tempTelegram.data[7];
                                                   #statReceive.configTelegramV2.lifeSignCycle := DWORD_TO_TIME(#tempDWord);
                                                   #diagnostics.partnerConfig.connnection.lifeSignCycleTime := #statReceive.configTelegramV2.lifeSignCycle;

                                                   //Sender cycleTime
                                                   #tempDWord.%B3 := #statReceive.tempTelegram.data[8];
                                                   #tempDWord.%B2 := #statReceive.tempTelegram.data[9];
                                                   #tempDWord.%B1 := #statReceive.tempTelegram.data[10];
                                                   #tempDWord.%B0 := #statReceive.tempTelegram.data[11];
                                                   #statReceive.configTelegramV2.cycleTime := DWORD_TO_TIME(#tempDWord);
                                                   #diagnostics.partnerConfig.sender.cycleTime := #statReceive.configTelegramV2.cycleTime;
                                                   //Sender ackTimeOut
                                                   #tempDWord.%B3 := #statReceive.tempTelegram.data[12];
                                                   #tempDWord.%B2 := #statReceive.tempTelegram.data[13];
                                                   #tempDWord.%B1 := #statReceive.tempTelegram.data[14];
                                                   #tempDWord.%B0 := #statReceive.tempTelegram.data[15];
                                                   #statReceive.configTelegramV2.ackTimeOut := DWORD_TO_TIME(#tempDWord);
                                                   #diagnostics.partnerConfig.sender.ackTimeout := #statReceive.configTelegramV2.ackTimeOut;
                                                   //MaxSendDataLength
                                                   #tempDWord.%B3 := #statReceive.tempTelegram.data[16];
                                                   #tempDWord.%B2 := #statReceive.tempTelegram.data[17];
                                                   #tempDWord.%B1 := #statReceive.tempTelegram.data[18];
                                                   #tempDWord.%B0 := #statReceive.tempTelegram.data[19];
                                                   #statReceive.configTelegramV2.maxSendDataLength := #tempDWord;
                                                   #diagnostics.partnerConfig.sizeOfSendBuffer := #statReceive.configTelegramV2.maxSendDataLength;
                                                   //MaxReceiveDataLength
                                                   #tempDWord.%B3 := #statReceive.tempTelegram.data[20];
                                                   #tempDWord.%B2 := #statReceive.tempTelegram.data[21];
                                                   #tempDWord.%B1 := #statReceive.tempTelegram.data[22];
                                                   #tempDWord.%B0 := #statReceive.tempTelegram.data[23];
                                                   #statReceive.configTelegramV2.maxReceiveDataLength := #tempDWord;
                                                   #diagnostics.partnerConfig.sizeOfReceiveBuffer := #statReceive.configTelegramV2.maxReceiveDataLength;

                                                   //Set FB.#connected and #diagnostics information
                                                   #connected := #statConnected := TRUE;
                                                   #diagnostics.statistics.LComProtocolUsed := TRUE;
                                                   #diagnostics.statistics.activeLComVersion := #HEADER_V2;
                                                   #statState.cfgSender := #OPERATION;

                                                   //Write diagnostics
                                                   #statDiag.bufferIndex := #statDiag.bufferIndex + 1;
                                                   #statDiag.buffer[#statDiag.bufferIndex].status := #STATUS_CONNECTED_V2;
                                                   #statDiag.buffer[#statDiag.bufferIndex].subFunctionErrorID := 16#0000;
                                                   #statDiag.buffer[#statDiag.bufferIndex].additionalValue1 := 0.0;
                                                   #statDiag.buffer[#statDiag.bufferIndex].additionalValue2 := 0.0;
                                                   #statDiag.buffer[#statDiag.bufferIndex].additionalValue3 := 0.0;
                                                   #statDiag.buffer[#statDiag.bufferIndex].additionalValue4 := T#0ms;

                                                   //Check timeSync setting at local cpu and partner cpu
                                                   IF ((#diagnostics.localConfig.timeSync.usePartnerTimestamps
                                                       XOR
                                                       #diagnostics.partnerConfig.timeSync.usePartnerTimestamps)
                                                       AND
                                                       (#diagnostics.localConfig.timeSync.sendMode > 0
                                                       OR
                                                       #diagnostics.partnerConfig.timeSync.sendMode > 0))
                                                   THEN
                                                       ;//One cpu does send timeSync information
                                                   ELSE
                                                       //Write diagnostics
                                                       #statDiag.bufferIndex := #statDiag.bufferIndex + 1;
                                                       #statDiag.buffer[#statDiag.bufferIndex].status := #WARN_NO_TIME_SYNC;
                                                       #statDiag.buffer[#statDiag.bufferIndex].subFunctionErrorID := 16#0000;
                                                       #statDiag.buffer[#statDiag.bufferIndex].additionalValue1 := 0.0;
                                                       #statDiag.buffer[#statDiag.bufferIndex].additionalValue2 := 0.0;
                                                       #statDiag.buffer[#statDiag.bufferIndex].additionalValue3 := 0.0;
                                                       #statDiag.buffer[#statDiag.bufferIndex].additionalValue4 := T#0ms;
                                                   END_IF;
                                                   //Do not send telegram 1
                                               ELSE
                                                   //LCom V1
                                                   //LifeSignCycle
                                                   #statReceive.configTelegramV1.lifeSignCycle.%B1 := #statReceive.tempTelegram.data[8];
                                                   #statReceive.configTelegramV1.lifeSignCycle.%B0 := #statReceive.tempTelegram.data[9];
                                                   #diagnostics.partnerConfig.connnection.lifeSignCycleTime := UINT_TO_TIME(#statReceive.configTelegramV1.lifeSignCycle);
                                                   //CycleTime
                                                   #statReceive.configTelegramV1.cycleTime.%B1 := #statReceive.tempTelegram.data[4];
                                                   #statReceive.configTelegramV1.cycleTime.%B0 := #statReceive.tempTelegram.data[5];
                                                   #diagnostics.partnerConfig.sender.cycleTime := UINT_TO_TIME(#statReceive.configTelegramV1.cycleTime);
                                                   //AckTimeOut
                                                   #statReceive.configTelegramV1.ackTimeOut.%B1 := #statReceive.tempTelegram.data[6];
                                                   #statReceive.configTelegramV1.ackTimeOut.%B0 := #statReceive.tempTelegram.data[7];
                                                   #diagnostics.partnerConfig.sender.ackTimeout := UINT_TO_TIME(#statReceive.configTelegramV1.ackTimeOut);
                                                   //MaxSendDataLength
                                                   #statReceive.configTelegramV1.maxSendDataLength.%B1 := #statReceive.tempTelegram.data[12];
                                                   #statReceive.configTelegramV1.maxSendDataLength.%B0 := #statReceive.tempTelegram.data[13];
                                                   #diagnostics.partnerConfig.sizeOfSendBuffer := #statReceive.configTelegramV1.maxSendDataLength;
                                                   //MaxReceiveDataLength
                                                   #statReceive.configTelegramV1.maxReceiveDataLength.%B1 := #statReceive.tempTelegram.data[14];
                                                   #statReceive.configTelegramV1.maxReceiveDataLength.%B0 := #statReceive.tempTelegram.data[15];
                                                   #diagnostics.partnerConfig.sizeOfReceiveBuffer := #statReceive.configTelegramV1.maxReceiveDataLength;
                                                   //UsesTimeStamp
                                                   #diagnostics.partnerConfig.timeSync.usePartnerTimestamps := BYTE_TO_BOOL(#statReceive.tempTelegram.data[10]);
                                                   //SendModeSyncTime
                                                   #diagnostics.partnerConfig.timeSync.sendMode := #statReceive.tempTelegram.data[11];

                                                   //Send Telegram 1
                                                   #statSend.tsendFct.data[#statSend.tsendFct.dataOffset] := #statSend.configTelegramV1.LComVersion;
                                                   #statSend.tsendFct.data[#statSend.tsendFct.dataOffset + 1] := 16#01;
                                                   #statSend.tsendFct.data[#statSend.tsendFct.dataOffset + 2] := #statSend.configTelegramV1.comMode;
                                                   #statSend.tsendFct.data[#statSend.tsendFct.dataOffset + 3] := #statSend.configTelegramV1.slidingWindow;
                                                   //CycleTime
                                                   #statSend.tsendFct.data[#statSend.tsendFct.dataOffset + 4] := #statReceive.configTelegramV1.cycleTime.%B1;
                                                   #statSend.tsendFct.data[#statSend.tsendFct.dataOffset + 5] := #statReceive.configTelegramV1.cycleTime.%B0;
                                                   //AckTimeOut
                                                   #statSend.tsendFct.data[#statSend.tsendFct.dataOffset + 6] := #statReceive.configTelegramV1.ackTimeOut.%B1;
                                                   #statSend.tsendFct.data[#statSend.tsendFct.dataOffset + 7] := #statReceive.configTelegramV1.ackTimeOut.%B0;
                                                   //LifeSignCycle
                                                   #statSend.tsendFct.data[#statSend.tsendFct.dataOffset + 8] := #statSend.configTelegramV1.lifeSignCycle.%B1;
                                                   #statSend.tsendFct.data[#statSend.tsendFct.dataOffset + 9] := #statSend.configTelegramV1.lifeSignCycle.%B0;
                                                   //Status
                                                   #statSend.tsendFct.data[#statSend.tsendFct.dataOffset + 10] := #statSend.configTelegramV1.status;
                                                   //SendModeSyncTime
                                                   #statSend.tsendFct.data[#statSend.tsendFct.dataOffset + 11] := #statSend.configTelegramV1.sendModeSyncTime;
                                                   //MaxSendDataLength
                                                   #statSend.tsendFct.data[#statSend.tsendFct.dataOffset + 12] := #statSend.configTelegramV1.maxSendDataLength.%B1;
                                                   #statSend.tsendFct.data[#statSend.tsendFct.dataOffset + 13] := #statSend.configTelegramV1.maxSendDataLength.%B0;
                                                   //MaxReceiveDataLength
                                                   #statSend.tsendFct.data[#statSend.tsendFct.dataOffset + 14] := #statSend.configTelegramV1.maxReceiveDataLength.%B1;
                                                   #statSend.tsendFct.data[#statSend.tsendFct.dataOffset + 15] := #statSend.configTelegramV1.maxReceiveDataLength.%B0;
                                                   //Calculate offset in the tcp send buffer
                                                   #statSend.tsendFct.dataOffset := #statSend.tsendFct.dataOffset + 16;
                                                   //Set state
                                                   #statState.sender := #SEND_CONFIG;
                                               END_IF;

                                           5://Telegram type 5

                                               //Reset index, so a new temp. LCom header can be built
                                               #statReceive.tempTelegram.index := 0;
                                               #statReceive.numberOfLComHeader := #statReceive.numberOfLComHeader + 1;

                                               //Accept timestamp from partner ?
                                               IF (#diagnostics.localConfig.timeSync.usePartnerTimestamps) THEN
                                                   //Yes --> Accept timestamp from partner
                                                   #tempActTime.YEAR := INT_TO_UINT(BCD16_TO_INT(#statReceive.tempTelegram.data[2] AND 16#00FF));
                                                   IF ((#tempActTime.YEAR >= 90)
                                                       AND (#tempActTime.YEAR <= 99))
                                                   THEN
                                                       #tempActTime.YEAR := #tempActTime.YEAR + 1900;
                                                   ELSE
                                                       #tempActTime.YEAR := #tempActTime.YEAR + 2000;
                                                   END_IF;

                                                   #tempActTime.MONTH := INT_TO_USINT(BCD16_TO_INT(#statReceive.tempTelegram.data[3] AND 16#00FF));
                                                   #tempActTime.DAY := INT_TO_USINT(BCD16_TO_INT(#statReceive.tempTelegram.data[4] AND 16#00FF));
                                                   #tempActTime.HOUR := INT_TO_USINT(BCD16_TO_INT(#statReceive.tempTelegram.data[5] AND 16#00FF));
                                                   #tempActTime.MINUTE := INT_TO_USINT(BCD16_TO_INT(#statReceive.tempTelegram.data[6] AND 16#00FF));
                                                   #tempActTime.SECOND := INT_TO_USINT(BCD16_TO_INT(#statReceive.tempTelegram.data[7] AND 16#00FF));
                                                   #tempActTime.NANOSECOND := INT_TO_UDINT(BCD16_TO_INT(#statReceive.tempTelegram.data[8] AND 16#00FF));
                                                   #tempActTime.NANOSECOND := #tempActTime.NANOSECOND * 1000;
                                                   #tempActTime.NANOSECOND := #tempActTime.NANOSECOND + 500;
                                                   #tempActTime.WEEKDAY := INT_TO_USINT(BCD16_TO_INT(#statReceive.tempTelegram.data[9] AND 16#000F));
                                                   //Write local time
                                                   #statRet := WR_LOC_T(LOCTIME := #tempActTime, DST := FALSE);
                                                   //Statistic --> Get time stamp of last time sync
                                                   #diagnostics.statistics.lastTimeSync := #tempActTime;
                                               ELSE
                                                   ;//No --> Do not write system time
                                               END_IF;

                                           20://Telegram type 20

                                               //Reset index, so a new temp. LCom header can be built
                                               #statReceive.numberOfLComHeader := #statReceive.numberOfLComHeader + 1;
                                               #statReceive.tempTelegram.index := 0;

                                               //Write diagnostics ---> Stop analyzing the tcp receive buffer
                                               #statDiag.bufferIndex := #statDiag.bufferIndex + 1;
                                               #statDiag.buffer[#statDiag.bufferIndex].status := #STATUS_DISCONNECTING;
                                               #statDiag.buffer[#statDiag.bufferIndex].subFunctionErrorID := 16#0000;
                                               #statDiag.buffer[#statDiag.bufferIndex].additionalValue1 := 0.0;
                                               #statDiag.buffer[#statDiag.bufferIndex].additionalValue2 := 0.0;
                                               #statDiag.buffer[#statDiag.bufferIndex].additionalValue3 := 0.0;
                                               #statDiag.buffer[#statDiag.bufferIndex].additionalValue4 := T#0ms;
                                               #statState.connection := #CLOSE_CONNECTION;
                                               EXIT;

                                           ELSE//Telegram type is unknown
                                               //Write diagnostics
                                               #statDiag.bufferIndex := #statDiag.bufferIndex + 1;
                                               #statDiag.buffer[#statDiag.bufferIndex].status := #ERR_WRONG_TELEGRAM_ID;
                                               #statDiag.buffer[#statDiag.bufferIndex].subFunctionErrorID := 16#0000;
                                               #statDiag.buffer[#statDiag.bufferIndex].additionalValue1 := #statReceive.tempTelegram.telegramType;
                                               #statDiag.buffer[#statDiag.bufferIndex].additionalValue2 := 0.0;
                                               #statDiag.buffer[#statDiag.bufferIndex].additionalValue3 := 0.0;
                                               #statDiag.buffer[#statDiag.bufferIndex].additionalValue4 := T#0ms;
                                               #statState.connection := #CLOSE_CONNECTION;
                                               GOTO diag;
                                       END_CASE;

                                   END_IF;
                               END_REGION LCOM_PROTOCOL

                               //Calculate rest of data in the tcp receive buffer
                               #statReceive.trcvFct.dataLengthRest := #statReceive.trcvFct.dataLength - #statReceive.trcvFct.dataOffset;

                           UNTIL ((#statReceive.trcvFct.dataLengthRest <= 0)
                               OR (#statReceive.trcvFct.dataLengthRest > #MAX_DATA_BUFFER))
                               //If the result of the calculation of the rest data is greater than 4096, then an error occurred
                           END_REPEAT;
                           //End:Analyze tcp receive buffer with LCom protocol

                       END_IF;//#readDataLength <> 0
                   END_REGION READ_TCP_BUFFER

                   REGION HANDLE_SENDING
                       //---------------------------------------------------------------------
                       //Check if next package can be sent
                       //---------------------------------------------------------------------
                       IF ((#statConnected = TRUE) AND (#statState.connection = #OPERATION)) THEN

                           //Get cycle time [ms]
                           #instLocalCycleTimeTimer(IN := TRUE,
                                                    PT := #diagnostics.localConfig.sender.cycleTime);


                           //---------------------------------------------------------------------
                           //In sending process
                           //---------------------------------------------------------------------
                           IF (#statSending = TRUE) THEN
                               //Yes --> In sending process

                               REGION CHECK_SEND_CYCLETIME
                                   //---------------------------------------------------------------------
                                   //Check if sender cycle time is expired (with and without LCom protocol) ?
                                   //---------------------------------------------------------------------
                                   IF (#instLocalCycleTimeTimer.Q AND #diagnostics.localConfig.sender.cycleTime > T#0ms) THEN
                                       //Yes --> Sender cycle time is expired
                                       //Check if sender cycle time violation is already stored ?
                                       IF (#statSend.userData.sendCycleViolation) THEN
                                           ;//Yes --> Exceeded before and stored
                                       ELSE
                                           //No --> Increase number of send cycle time violations
                                           #diagnostics.statistics.totalSendCycleViolations := #diagnostics.statistics.totalSendCycleViolations + 1;
                                           #statSend.userData.sendCycleViolation := TRUE;
                                       END_IF;

                                       //Write diagnostics
                                       #statDiag.bufferIndex := #statDiag.bufferIndex + 1;
                                       #statDiag.buffer[#statDiag.bufferIndex].status := #WARN_SEND_CYCLE_EXPIRED;
                                       #statDiag.buffer[#statDiag.bufferIndex].subFunctionErrorID := 16#0000;
                                       #statDiag.buffer[#statDiag.bufferIndex].additionalValue1 := UDINT_TO_REAL(TIME_TO_UDINT(#diagnostics.localConfig.sender.cycleTime));
                                       #statDiag.buffer[#statDiag.bufferIndex].additionalValue2 := 0.0;
                                       #statDiag.buffer[#statDiag.bufferIndex].additionalValue3 := 0.0;
                                       #statDiag.buffer[#statDiag.bufferIndex].additionalValue4 := #instLocalCycleTimeTimer.ET;
                                   ELSE
                                       ;//No --> Sender cycle time is not expired
                                   END_IF;//End: Check if sender cycle time is expired (with and without LCom protocol) ?
                               END_REGION CHECK_SEND_CYCLETIME

                               REGION CHECK_ACK_TIMEOUT
                                   //---------------------------------------------------------------------
                                   //Check acknowledge timeout with LCom protocol
                                   //---------------------------------------------------------------------
                                   IF (#diagnostics.localConfig.connection.useLComProtocol = TRUE) THEN

                                       //Get acknowledge timeout [ms]
                                       #instExpectedAckPackage1(IN := TRUE,
                                                                PT := #diagnostics.localConfig.sender.ackTimeout);

                                       //Check if acknowledge timeout is expired ?
                                       IF ((#instExpectedAckPackage1.Q = TRUE)
                                           AND
                                           (#statSend.numberOfLComPackage > 0))
                                       THEN
                                           //Yes --> Acknowledge timeout is expired, increase number of confirmation timeouts
                                           #diagnostics.statistics.totalAckTimeouts := #diagnostics.statistics.totalAckTimeouts + 1;

                                           //Write diagnostics
                                           #statDiag.bufferIndex := #statDiag.bufferIndex + 1;
                                           #statDiag.buffer[#statDiag.bufferIndex].status := #ERR_ACK_TIMEOUT_EXPIRED;
                                           #statDiag.buffer[#statDiag.bufferIndex].subFunctionErrorID := 16#0000;
                                           #statDiag.buffer[#statDiag.bufferIndex].additionalValue1 := UDINT_TO_REAL(TIME_TO_UDINT(#diagnostics.localConfig.sender.ackTimeout));
                                           #statDiag.buffer[#statDiag.bufferIndex].additionalValue2 := 0.0;
                                           #statDiag.buffer[#statDiag.bufferIndex].additionalValue3 := 0.0;
                                           #statDiag.buffer[#statDiag.bufferIndex].additionalValue4 := #instExpectedAckPackage1.ET;
                                           #statState.connection := #CLOSE_CONNECTION;
                                           GOTO diag;
                                       ELSE
                                           //No --> Acknowledge timeout is not expired

                                           //Is the last LCom package already sent ?
                                           IF (#statState.comSender = #SEND_NO_DATA) THEN
                                               ;//Yes --> Wait for acknowledge telegram
                                           ELSE
                                               //No --> Last LCom package not sent yet

                                               //Check if the next LCom package can be sent ? (Sliding window)
                                               IF ((#statSend.numberOfLComPackage < 1)
                                                   AND
                                                   (#diagnostics.statistics.activeLComVersion = #HEADER_V1
                                                   OR
                                                   #diagnostics.statistics.activeLComVersion = #HEADER_V2))
                                               THEN
                                                   //Yes --> Continue sending
                                                   #statState.comSender := #CYCLE;
                                               ELSE
                                                   //No --> Wait for acknowledge telegram
                                                   #statState.comSender := #WAIT_ACK_TELEGRAM;
                                               END_IF;
                                           END_IF;//End: Is the last LCom package already sent ?
                                       END_IF;//End: Check if acknowledge time is expired ?
                                   ELSE
                                       //Continue without LCom protocol, acknowledge timeout is not valid
                                       #statState.comSender := #CYCLE;
                                   END_IF;
                               END_REGION CHECK_ACK_TIMEOUT

                           ELSE
                               //Not --> Not in sending process
                               REGION CHECK_SEND_CONFIG_AND_DATA_TO_SEND
                                   //With LCom protocol --> Check if sender configuration was changed
                                   IF (#diagnostics.localConfig.connection.useLComProtocol = TRUE
                                       AND
                                       ((#configuration.sender.cycleTime <> #statCompare.sender.cycleTime)
                                       OR
                                       (#configuration.sender.ackTimeout <> #statCompare.sender.ackTimeOut)))
                                   THEN
                                       #connected := #statConnected := FALSE;
                                       //Update parameters
                                       #statState.cfgSender := #STATE_INIT;
                                   ELSIF (NOT #diagnostics.localConfig.connection.useLComProtocol
                                       AND
                                       #configuration.sender.cycleTime <> #statCompare.sender.cycleTime)
                                   THEN//Without LCom protocol --> Check if sender configuration was changed
                                       //Update parameters
                                       #diagnostics.localConfig.sender.cycleTime := #configuration.sender.cycleTime;
                                       #statCompare.sender.cycleTime := #configuration.sender.cycleTime;
                                   ELSIF (#send OR #statRisingEdgeSend)//Check if FB.send input is true or rising edge is detected ?
                                   THEN
                                       //Yes --> FB.send input is true

                                       //---------------------------------------------------------------------
                                       //Check if data have to be sent
                                       //---------------------------------------------------------------------
                                       IF ((#sendDataLength > 0)
                                           AND
                                           ((#statRisingEdgeSend)//Rising edge
                                           OR
                                           ((#instLocalCycleTimeTimer.Q)//check CycleTimeTimer
                                           AND
                                           (#diagnostics.localConfig.sender.cycleTime > T#0ms))))
                                       THEN
                                           //Start sending
                                           #sending := #statSending := TRUE;
                                           #statSend.userData.sendCycleViolation := FALSE;
                                           #statSend.userData.offset := 0;
                                           #statRisingEdgeSend := FALSE;

                                           //Start message sending timer
                                           #instMsgSendingTimer(IN := TRUE,
                                                                PT := T#+24d20h31m23s647ms);

                                           //Stop/Start local cycle timer
                                           #instLocalCycleTimeTimer(IN := FALSE,
                                                                    PT := #diagnostics.localConfig.sender.cycleTime);
                                           #instLocalCycleTimeTimer(IN := TRUE,
                                                                    PT := #diagnostics.localConfig.sender.cycleTime);


